FUNCTION_BLOCK "naut_Loop"
{ S7_Optimized_Access := 'TRUE' }
VERSION : 0.1
   VAR_INPUT
      Enable : BOOL;
      Meas : REAL;
      Target : REAL;
   END_VAR
   VAR_OUTPUT
      Out : REAL;
   END_VAR
   VAR
      ctl : "naut_PID";
   END_VAR

BEGIN
	#ctl(AUTO := #Enable, PV := #Meas, SP := #Target, KP := 2.0, KI := 0.5, CV_MIN := 0.0, CV_MAX := 100.0);
	#Out := #ctl.CV;
END_FUNCTION_BLOCK
